Fanuc KAREL source: KO00103.KL

PROGRAM KO00103
%NOLOCKGROUP
VAR
  A: INTEGER
  B: ARRAY[2] OF SHORT
  OUT: INTEGER
BEGIN
  A = 1
  B[1] = 2
  OUT = ATAN2(A, B[1])
END KO00103
